// TIA Portal V17 export
// export: Created 2026-11-10T15:00:48.6641979Z, ExportSetting WithDefaults, DisplayName Totally Integrated Automation Portal, DisplayVersion V17, DisplayName TIA Portal Openness, DisplayVersion V17, DisplayName TIA Portal Version Control Interface, DisplayVersion V17, DisplayName STEP 7 Professional, DisplayVersion V17, DisplayName STEP 7 Safety, DisplayVersion V17, DisplayName WinCC Advanced, DisplayVersion V17
GraphicList "Gauge120"  ListRange=Decimal, Mode=Simple
  GraphicListEntry   EntryType=Range, To=11, Picture=Gauge_0
  GraphicListEntry   EntryType=Range, From=12, To=23, Picture=Gauge_1
  GraphicListEntry   EntryType=Range, From=24, To=35, Picture=Gauge_2
  GraphicListEntry   EntryType=Range, From=36, To=47, Picture=Gauge_3
  GraphicListEntry   EntryType=Range, From=48, To=59, Picture=Gauge_4
  GraphicListEntry   EntryType=Range, From=60, To=71, Picture=Gauge_5
  GraphicListEntry   EntryType=Range, From=72, To=83, Picture=Gauge_6
  GraphicListEntry   EntryType=Range, From=84, To=95, Picture=Gauge_7
  GraphicListEntry   EntryType=Range, From=96, To=107, Picture=Gauge_8
  GraphicListEntry   EntryType=Range, From=108, To=119, Picture=Gauge_9
  GraphicListEntry   EntryType=Range, From=120, To=120, Picture=Gauge_10
